// TIA Portal V20 export
// export: Created 2026-10-30T08:30:38.2615563Z, ExportSetting WithDefaults, DisplayName Totally Integrated Automation Portal, DisplayVersion V20, DisplayName TIA Portal Openness, DisplayVersion V20, DisplayName TIA Portal Version Control Interface, DisplayVersion V20, DisplayName SIRIUS Safety ES, DisplayVersion V20, DisplayName STEP 7 Professional, DisplayVersion V20, DisplayName STEP 7 Safety, DisplayVersion V20, DisplayName WinCC Basic/Comfort/Advanced, DisplayVersion V20, DisplayName WinCC Professional, DisplayVersion V20, DisplayName WinCC Unified, DisplayVersion V20
FUNCTION "Block_1" : Void   // FC1, LAD
{ S7_Optimized_Access := 'TRUE' }
VERSION : 0.1
// stored: AutoNumber true, IsIECCheckEnabled false, SetENOAutomatically false, UDAEnableTagReadback false
BEGIN

REGION Network 1
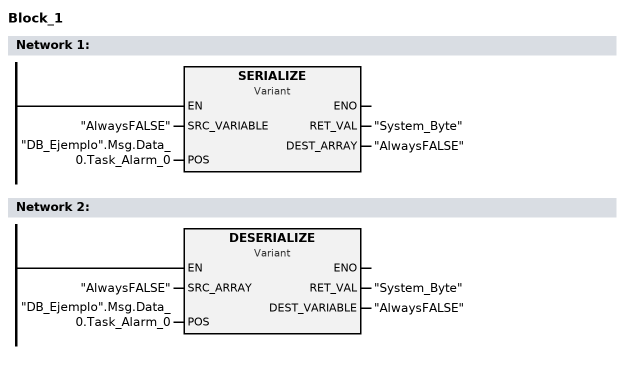
   RUNG wire#powerrail
      { S7_Templates := "[src_type := Variant, dest_type := Variant]" } Serialize(SRC_VARIABLE := "AlwaysFALSE", POS := "DB_Ejemplo".Msg.Data_0.Task_Alarm_0, Ret_Val => "System_Byte", DEST_ARRAY => "AlwaysFALSE")
   END_RUNG
   // the same network as SCL:
   "System_Byte" := Serialize(SRC_VARIABLE := "AlwaysFALSE",
                           POS := "DB_Ejemplo".Msg.Data_0.Task_Alarm_0,
                           DEST_ARRAY => "AlwaysFALSE");
END_REGION

REGION Network 2
   RUNG wire#powerrail
      { S7_Templates := "[src_type := Variant, dest_type := Variant]" } Deserialize(SRC_ARRAY := "AlwaysFALSE", POS := "DB_Ejemplo".Msg.Data_0.Task_Alarm_0, Ret_Val => "System_Byte", DEST_VARIABLE => "AlwaysFALSE")
   END_RUNG
   // the same network as SCL:
   "System_Byte" := Deserialize(SRC_ARRAY := "AlwaysFALSE",
                           POS := "DB_Ejemplo".Msg.Data_0.Task_Alarm_0,
                           DEST_VARIABLE => "AlwaysFALSE");
END_REGION
END_FUNCTION
